Fanuc KAREL source: kt00447.KL

-- PROVISIONAL review KL for V1013-1; original PC SHA256 314f95aa091da0393de520ffa4e8d1cfc3d7bb279cc11d2b1f32d3714f040ffc
-- Incomplete behavior may be omitted. Consult companion uncertainty JSON. Do not deploy.
PROGRAM KT00447
%NOLOCKGROUP
VAR
  I2 : INTEGER
  OUT : BOOLEAN
-- UNRESOLVED_DECL Y1 type=002018
BEGIN
  -- UNRESOLVED_PC offsets 5-19; opcodes 2E,22,9D,33,B2
  -- UNRESOLVED_PC offsets 24-35; opcodes 2E,23
  -- UNRESOLVED_PC offsets 40-62; opcodes 22,9D,33,B1,21,5C,23
  -- UNRESOLVED_PC offsets 67-71; opcodes 7F
END KT00447
